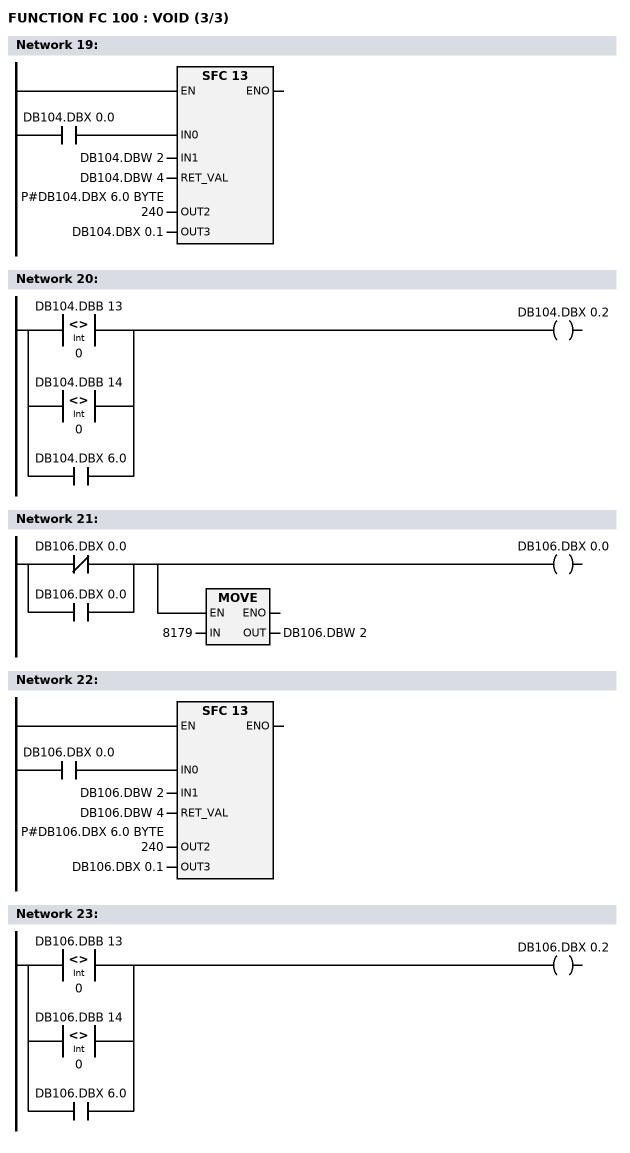

      A     DB104.DBX    0.0;
      =     L      0.0;
      BLD   103;
      CALL SFC   13 (
           IN0                      := L      0.0,
           IN1                      := DB104.DBW    2,
           RET_VAL                  := DB104.DBW    4,
           OUT2                     := P#DB104.DBX 6.0 BYTE 240,
           OUT3                     := DB104.DBX    0.1);
      NOP   0;
NETWORK
TITLE =

      O(    ;
      L     DB104.DBB   13;
      L     0;
      <>I   ;
      )     ;
      O(    ;
      L     DB104.DBB   14;
      L     0;
      <>I   ;
      )     ;
      O     DB104.DBX    6.0;
      =     DB104.DBX    0.2;
NETWORK
TITLE =

      ON    DB106.DBX    0.0;
      O     DB106.DBX    0.0;
      =     L      0.0;
      A     L      0.0;
      BLD   102;
      =     DB106.DBX    0.0;
      A     L      0.0;
      JNB   M003;
      L     8179;
      T     DB106.DBW    2;
M003: NOP   0;
NETWORK
TITLE =

      A     DB106.DBX    0.0;
      =     L      0.0;
      BLD   103;
      CALL SFC   13 (
           IN0                      := L      0.0,
           IN1                      := DB106.DBW    2,
           RET_VAL                  := DB106.DBW    4,
           OUT2                     := P#DB106.DBX 6.0 BYTE 240,
           OUT3                     := DB106.DBX    0.1);
      NOP   0;
NETWORK
TITLE =

      O(    ;
      L     DB106.DBB   13;
      L     0;
      <>I   ;
      )     ;
      O(    ;
      L     DB106.DBB   14;
      L     0;
      <>I   ;
      )     ;
      O     DB106.DBX    6.0;
      =     DB106.DBX    0.2;
END_FUNCTION

DATA_BLOCK DB 500
VERSION : 0.0

 FB 500
BEGIN
   IN0 := FALSE;
   IN1 := FALSE;
   IN2 := FALSE;
   OUT3 := FALSE;
   OUT4 := FALSE;
   STAT5 := FALSE;
   STAT6 := FALSE;
   STAT7 := FALSE;
   STAT8 := FALSE;
END_DATA_BLOCK

DATA_BLOCK DB 501
VERSION : 0.0

 FB 500
BEGIN
   IN0 := FALSE;
   IN1 := FALSE;
   IN2 := FALSE;
   OUT3 := FALSE;
   OUT4 := FALSE;
   STAT5 := FALSE;
   STAT6 := FALSE;
   STAT7 := FALSE;
   STAT8 := FALSE;
END_DATA_BLOCK

DATA_BLOCK DB 502
VERSION : 0.0

 FB 500
BEGIN
   IN0 := FALSE;
   IN1 := FALSE;
   IN2 := FALSE;
   OUT3 := FALSE;
   OUT4 := FALSE;
   STAT5 := FALSE;
   STAT6 := FALSE;
   STAT7 := FALSE;
   STAT8 := FALSE;
END_DATA_BLOCK

DATA_BLOCK DB 504
VERSION : 0.0

 FB 500
BEGIN
   IN0 := FALSE;
   IN1 := FALSE;
   IN2 := FALSE;
   OUT3 := FALSE;
   OUT4 := FALSE;
   STAT5 := FALSE;
   STAT6 := FALSE;
   STAT7 := FALSE;
   STAT8 := FALSE;
END_DATA_BLOCK

DATA_BLOCK DB 505
VERSION : 0.0

 FB 500
BEGIN
   IN0 := FALSE;
   IN1 := FALSE;
   IN2 := FALSE;
   OUT3 := FALSE;
   OUT4 := FALSE;
   STAT5 := FALSE;
   STAT6 := FALSE;
   STAT7 := FALSE;
   STAT8 := FALSE;
END_DATA_BLOCK

DATA_BLOCK DB 506
VERSION : 0.0

 FB 500
BEGIN
   IN0 := FALSE;
   IN1 := FALSE;
   IN2 := FALSE;
   OUT3 := FALSE;
   OUT4 := FALSE;
   STAT5 := FALSE;
   STAT6 := FALSE;
   STAT7 := FALSE;
   STAT8 := FALSE;
END_DATA_BLOCK

DATA_BLOCK DB 507
VERSION : 0.0

 FB 500
BEGIN
   IN0 := FALSE;
   IN1 := FALSE;
   IN2 := FALSE;
   OUT3 := FALSE;
   OUT4 := FALSE;
   STAT5 := FALSE;
   STAT6 := FALSE;
   STAT7 := FALSE;
   STAT8 := FALSE;
END_DATA_BLOCK

DATA_BLOCK DB 508
VERSION : 0.0

 FB 500
BEGIN
   IN0 := FALSE;
   IN1 := FALSE;
   IN2 := FALSE;
   OUT3 := FALSE;
   OUT4 := FALSE;
   STAT5 := FALSE;
   STAT6 := FALSE;
   STAT7 := FALSE;
   STAT8 := FALSE;
END_DATA_BLOCK

DATA_BLOCK DB 509
VERSION : 0.0

 FB 500
BEGIN
   IN0 := FALSE;
   IN1 := FALSE;
   IN2 := FALSE;
   OUT3 := FALSE;
   OUT4 := FALSE;
   STAT5 := FALSE;
   STAT6 := FALSE;
   STAT7 := FALSE;
   STAT8 := FALSE;
END_DATA_BLOCK

DATA_BLOCK DB 512
VERSION : 0.0

 FB 500
BEGIN
   IN0 := FALSE;
   IN1 := FALSE;
   IN2 := FALSE;
   OUT3 := FALSE;
   OUT4 := FALSE;
   STAT5 := FALSE;
   STAT6 := FALSE;
   STAT7 := FALSE;
   STAT8 := FALSE;
END_DATA_BLOCK

DATA_BLOCK DB 516
VERSION : 0.0

 FB 500
BEGIN
   IN0 := FALSE;
   IN1 := FALSE;
   IN2 := FALSE;
   OUT3 := FALSE;
   OUT4 := FALSE;
   STAT5 := FALSE;
   STAT6 := FALSE;
   STAT7 := FALSE;
   STAT8 := FALSE;
END_DATA_BLOCK

DATA_BLOCK DB 517
VERSION : 0.0

 FB 500
BEGIN
   IN0 := FALSE;
   IN1 := FALSE;
   IN2 := FALSE;
   OUT3 := FALSE;
   OUT4 := FALSE;
   STAT5 := FALSE;
   STAT6 := FALSE;
   STAT7 := FALSE;
   STAT8 := FALSE;
END_DATA_BLOCK

DATA_BLOCK DB 518
VERSION : 0.0

 FB 500
BEGIN
   IN0 := FALSE;
   IN1 := FALSE;
   IN2 := FALSE;
   OUT3 := FALSE;
   OUT4 := FALSE;
   STAT5 := FALSE;
   STAT6 := FALSE;
   STAT7 := FALSE;
   STAT8 := FALSE;
END_DATA_BLOCK

DATA_BLOCK DB 520
VERSION : 0.0

 FB 500
BEGIN
   IN0 := FALSE;
   IN1 := FALSE;
   IN2 := FALSE;
   OUT3 := FALSE;
   OUT4 := FALSE;
   STAT5 := FALSE;
   STAT6 := FALSE;
   STAT7 := FALSE;
   STAT8 := FALSE;
END_DATA_BLOCK

DATA_BLOCK DB 521
VERSION : 0.0

 FB 500
BEGIN
   IN0 := FALSE;
   IN1 := FALSE;
   IN2 := FALSE;
   OUT3 := FALSE;
   OUT4 := FALSE;
   STAT5 := FALSE;
   STAT6 := FALSE;
   STAT7 := FALSE;
   STAT8 := FALSE;
END_DATA_BLOCK

DATA_BLOCK DB 522
VERSION : 0.0

 FB 500
BEGIN
   IN0 := FALSE;
   IN1 := FALSE;
   IN2 := FALSE;
   OUT3 := FALSE;
   OUT4 := FALSE;
   STAT5 := FALSE;
   STAT6 := FALSE;
   STAT7 := FALSE;
   STAT8 := FALSE;
END_DATA_BLOCK

DATA_BLOCK DB 523
VERSION : 0.0

 FB 500
BEGIN
   IN0 := FALSE;
   IN1 := FALSE;
   IN2 := FALSE;
   OUT3 := FALSE;
   OUT4 := FALSE;
   STAT5 := FALSE;
   STAT6 := FALSE;
   STAT7 := FALSE;
   STAT8 := FALSE;
END_DATA_BLOCK

DATA_BLOCK DB 525
VERSION : 0.0

 FB 500
BEGIN
   IN0 := FALSE;
   IN1 := FALSE;
   IN2 := FALSE;
   OUT3 := FALSE;
   OUT4 := FALSE;
   STAT5 := FALSE;
   STAT6 := FALSE;
   STAT7 := FALSE;
   STAT8 := FALSE;
END_DATA_BLOCK

DATA_BLOCK DB 526
VERSION : 0.0

 FB 500
BEGIN
   IN0 := FALSE;
   IN1 := FALSE;
   IN2 := FALSE;
   OUT3 := FALSE;
   OUT4 := FALSE;
   STAT5 := FALSE;
   STAT6 := FALSE;
   STAT7 := FALSE;
   STAT8 := FALSE;
END_DATA_BLOCK

DATA_BLOCK DB 527
VERSION : 0.0

 FB 500
BEGIN
   IN0 := FALSE;
   IN1 := FALSE;
   IN2 := FALSE;
   OUT3 := FALSE;
   OUT4 := FALSE;
   STAT5 := FALSE;
   STAT6 := FALSE;
   STAT7 := FALSE;
   STAT8 := FALSE;
END_DATA_BLOCK

DATA_BLOCK DB 528
VERSION : 0.0

 FB 500
BEGIN
   IN0 := FALSE;
   IN1 := FALSE;
   IN2 := FALSE;
   OUT3 := FALSE;
   OUT4 := FALSE;
   STAT5 := FALSE;
   STAT6 := FALSE;
   STAT7 := FALSE;
   STAT8 := FALSE;
END_DATA_BLOCK

DATA_BLOCK DB 529
VERSION : 0.0

 FB 500
BEGIN
   IN0 := FALSE;
   IN1 := FALSE;
   IN2 := FALSE;
   OUT3 := FALSE;
   OUT4 := FALSE;
   STAT5 := FALSE;
   STAT6 := FALSE;
   STAT7 := FALSE;
   STAT8 := FALSE;
END_DATA_BLOCK

DATA_BLOCK DB 530
VERSION : 0.0

 FB 500
BEGIN
   IN0 := FALSE;
   IN1 := FALSE;
   IN2 := FALSE;
   OUT3 := FALSE;
   OUT4 := FALSE;
   STAT5 := FALSE;
   STAT6 := FALSE;
   STAT7 := FALSE;
   STAT8 := FALSE;
END_DATA_BLOCK

DATA_BLOCK DB 531
VERSION : 0.0

 FB 500
BEGIN
   IN0 := FALSE;
   IN1 := FALSE;
   IN2 := FALSE;
   OUT3 := FALSE;
   OUT4 := FALSE;
   STAT5 := FALSE;
   STAT6 := FALSE;
   STAT7 := FALSE;
   STAT8 := FALSE;
END_DATA_BLOCK

DATA_BLOCK DB 532
VERSION : 0.0

 FB 500
BEGIN
   IN0 := FALSE;
   IN1 := FALSE;
   IN2 := FALSE;
   OUT3 := FALSE;
   OUT4 := FALSE;
   STAT5 := FALSE;
   STAT6 := FALSE;
   STAT7 := FALSE;
   STAT8 := FALSE;
END_DATA_BLOCK

DATA_BLOCK DB 534
VERSION : 0.0

 FB 500
BEGIN
   IN0 := FALSE;
   IN1 := FALSE;
   IN2 := FALSE;
   OUT3 := FALSE;
   OUT4 := FALSE;
   STAT5 := FALSE;
   STAT6 := FALSE;
   STAT7 := FALSE;
   STAT8 := FALSE;
END_DATA_BLOCK

DATA_BLOCK DB 535
VERSION : 0.0

 FB 500
BEGIN
   IN0 := FALSE;
   IN1 := FALSE;
   IN2 := FALSE;
   OUT3 := FALSE;
   OUT4 := FALSE;
   STAT5 := FALSE;
   STAT6 := FALSE;
   STAT7 := FALSE;
   STAT8 := FALSE;
END_DATA_BLOCK

DATA_BLOCK DB 510
VERSION : 0.0

 FB 500
BEGIN
   IN0 := FALSE;
   IN1 := FALSE;
   IN2 := FALSE;
   OUT3 := FALSE;
   OUT4 := FALSE;
   STAT5 := FALSE;
   STAT6 := FALSE;
   STAT7 := FALSE;
   STAT8 := FALSE;
END_DATA_BLOCK

DATA_BLOCK DB 511
VERSION : 0.0

 FB 500
BEGIN
   IN0 := FALSE;
   IN1 := FALSE;
   IN2 := FALSE;
   OUT3 := FALSE;
   OUT4 := FALSE;
   STAT5 := FALSE;
   STAT6 := FALSE;
   STAT7 := FALSE;
   STAT8 := FALSE;
END_DATA_BLOCK

DATA_BLOCK DB 513
VERSION : 0.0

 FB 500
BEGIN
   IN0 := FALSE;
   IN1 := FALSE;
   IN2 := FALSE;
   OUT3 := FALSE;
   OUT4 := FALSE;
   STAT5 := FALSE;
   STAT6 := FALSE;
   STAT7 := FALSE;
   STAT8 := FALSE;
END_DATA_BLOCK

DATA_BLOCK DB 514
VERSION : 0.0

 FB 500
BEGIN
   IN0 := FALSE;
   IN1 := FALSE;
   IN2 := FALSE;
   OUT3 := FALSE;
   OUT4 := FALSE;
   STAT5 := FALSE;
   STAT6 := FALSE;
   STAT7 := FALSE;
   STAT8 := FALSE;
END_DATA_BLOCK

DATA_BLOCK DB 515
VERSION : 0.0

 FB 500
BEGIN
   IN0 := FALSE;
   IN1 := FALSE;
   IN2 := FALSE;
   OUT3 := FALSE;
   OUT4 := FALSE;
   STAT5 := FALSE;
   STAT6 := FALSE;
   STAT7 := FALSE;
   STAT8 := FALSE;
END_DATA_BLOCK

DATA_BLOCK DB 519
VERSION : 0.0

 FB 500
BEGIN
   IN0 := FALSE;
   IN1 := FALSE;
   IN2 := FALSE;
   OUT3 := FALSE;
   OUT4 := FALSE;
   STAT5 := FALSE;
   STAT6 := FALSE;
   STAT7 := FALSE;
   STAT8 := FALSE;
END_DATA_BLOCK

DATA_BLOCK DB 524
VERSION : 0.0

 FB 500
BEGIN
   IN0 := FALSE;
   IN1 := FALSE;
   IN2 := FALSE;
   OUT3 := FALSE;
   OUT4 := FALSE;
   STAT5 := FALSE;
   STAT6 := FALSE;
   STAT7 := FALSE;
   STAT8 := FALSE;
END_DATA_BLOCK

DATA_BLOCK DB 533
VERSION : 0.0

 FB 500
BEGIN
   IN0 := FALSE;
   IN1 := FALSE;
   IN2 := FALSE;
   OUT3 := FALSE;
   OUT4 := FALSE;
   STAT5 := FALSE;
   STAT6 := FALSE;
   STAT7 := FALSE;
   STAT8 := FALSE;
END_DATA_BLOCK

ORGANIZATION_BLOCK OB 1
VERSION : 0.1


VAR_TEMP
  TEMP0 : BYTE ;
  TEMP1 : BYTE ;
  TEMP2 : BYTE ;
  TEMP3 : BYTE ;
  TEMP4 : BYTE ;
  TEMP5 : BYTE ;
  TEMP6 : INT ;
  TEMP7 : INT ;
  TEMP8 : INT ;
  TEMP9 : DATE_AND_TIME ;
END_VAR
BEGIN
NETWORK
TITLE =
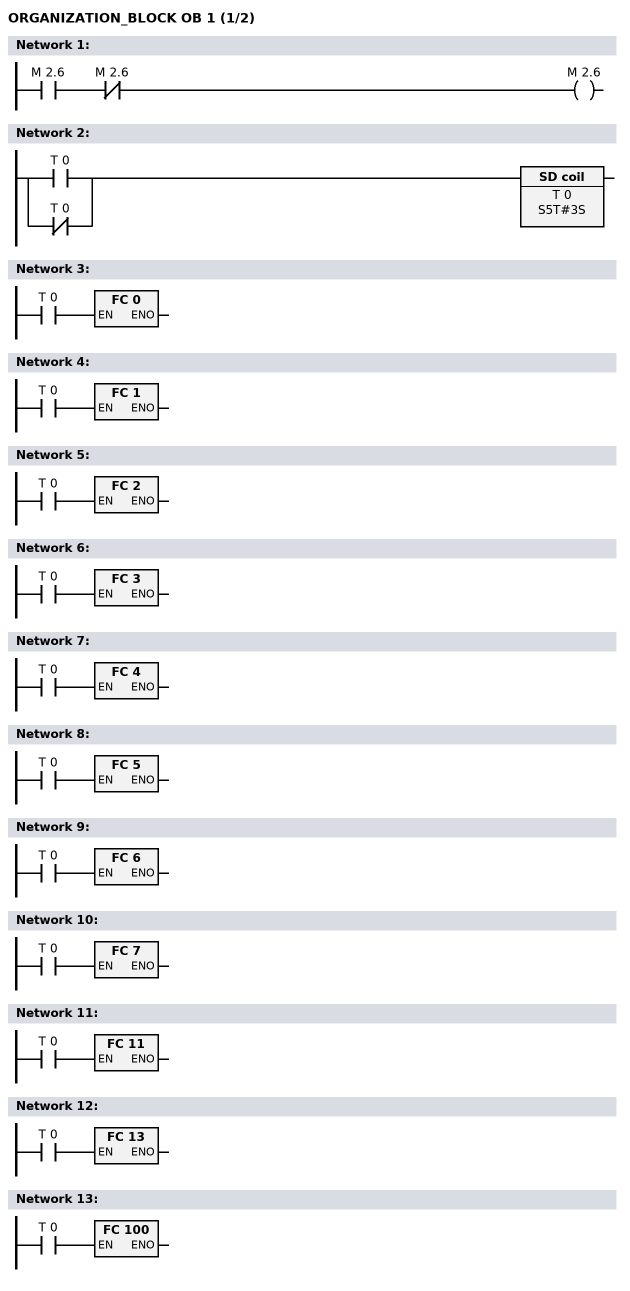

      A     M      2.6;
      AN    M      2.6;
      =     M      2.6;
NETWORK
TITLE =

      A(    ;
      O     T      0;
      ON    T      0;
      )     ;
      L     S5T#3S;
      SD    T      0;
      NOP   0;
      NOP   0;
      NOP   0;
      NOP   0;
NETWORK
TITLE =

      A     T      0;
      JNB   M001;
      CALL FC     0 ;
M001: NOP   0;
NETWORK
TITLE =

      A     T      0;
      JNB   M002;
      CALL FC     1 ;
M002: NOP   0;
NETWORK
TITLE =

      A     T      0;
      JNB   M003;
      CALL FC     2 ;
M003: NOP   0;
NETWORK
TITLE =

      A     T      0;
      JNB   M004;
      CALL FC     3 ;
M004: NOP   0;
NETWORK
TITLE =

      A     T      0;
      JNB   M005;
      CALL FC     4 ;
M005: NOP   0;
NETWORK
TITLE =

      A     T      0;
      JNB   M006;
      CALL FC     5 ;
M006: NOP   0;
NETWORK
TITLE =

      A     T      0;
      JNB   M007;
      CALL FC     6 ;
M007: NOP   0;
NETWORK
TITLE =

      A     T      0;
      JNB   M008;
      CALL FC     7 ;
M008: NOP   0;
NETWORK
TITLE =

      A     T      0;
      JNB   M009;
      CALL FC    11 ;
M009: NOP   0;
NETWORK
TITLE =

      A     T      0;
      JNB   M00a;
      CALL FC    13 ;
M00a: NOP   0;
NETWORK
TITLE =

      A     T      0;
      JNB   M00b;
      CALL FC   100 ;
M00b: NOP   0;
NETWORK
TITLE =
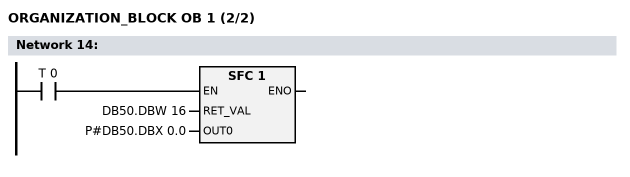

      A     T      0;
      JNB   M00c;
      CALL SFC    1 (
           RET_VAL                  := DB50.DBW   16,
           OUT0                     := P#DB50.DBX 0.0);
M00c: NOP   0;
END_ORGANIZATION_BLOCK

ORGANIZATION_BLOCK OB 35
VERSION : 0.1


VAR_TEMP
  TEMP0 : BYTE ;
  TEMP1 : BYTE ;
  TEMP2 : BYTE ;
  TEMP3 : BYTE ;
  TEMP4 : BYTE ;
  TEMP5 : BYTE ;
  TEMP6 : WORD ;
  TEMP7 : INT ;
  TEMP8 : INT ;
  TEMP9 : DATE_AND_TIME ;
END_VAR
BEGIN
END_ORGANIZATION_BLOCK

ORGANIZATION_BLOCK OB 70
VERSION : 0.1


VAR_TEMP
  TEMP0 : BYTE ;
  TEMP1 : BYTE ;
  TEMP2 : BYTE ;
  TEMP3 : BYTE ;
  TEMP4 : WORD ;
  TEMP5 : WORD ;
  TEMP6 : WORD ;
  TEMP7 : WORD ;
  TEMP8 : DATE_AND_TIME ;
END_VAR
BEGIN
NETWORK
TITLE =

      AN    M      3.7;
      =     M      3.7;
END_ORGANIZATION_BLOCK

ORGANIZATION_BLOCK OB 72
VERSION : 0.1


VAR_TEMP
  TEMP0 : BYTE ;
  TEMP1 : BYTE ;
  TEMP2 : BYTE ;
  TEMP3 : BYTE ;
  TEMP4 : WORD ;
  TEMP5 : WORD ;
  TEMP6 : WORD ;
  TEMP7 : WORD ;
  TEMP8 : DATE_AND_TIME ;
END_VAR
BEGIN
NETWORK
TITLE =

      A     M      3.7;
      =     M      3.7;
END_ORGANIZATION_BLOCK

ORGANIZATION_BLOCK OB 81
VERSION : 0.1


VAR_TEMP
  TEMP0 : BYTE ;
  TEMP1 : BYTE ;
  TEMP2 : BYTE ;
  TEMP3 : BYTE ;
  TEMP4 : BYTE ;
  TEMP5 : BYTE ;
  TEMP6 : WORD ;
  TEMP7 : BYTE ;
  TEMP8 : BYTE ;
  TEMP9 : BYTE ;
  TEMP10 : BYTE ;
  TEMP11 : DATE_AND_TIME ;
END_VAR
BEGIN
NETWORK
TITLE =

      AN    M      3.7;
      =     M      3.7;
END_ORGANIZATION_BLOCK

ORGANIZATION_BLOCK OB 82
VERSION : 0.1


VAR_TEMP
  TEMP0 : BYTE ;
  TEMP1 : BYTE ;
  TEMP2 : BYTE ;
  TEMP3 : BYTE ;
  TEMP4 : BYTE ;
  TEMP5 : BYTE ;
  TEMP6 : WORD ;
  TEMP7 : BOOL ;
  TEMP8 : BOOL ;
  TEMP9 : BOOL ;
  TEMP10 : BOOL ;
  TEMP11 : BOOL ;
  TEMP12 : BOOL ;
  TEMP13 : BOOL ;
  TEMP14 : BOOL ;
  TEMP15 : BYTE ;
  TEMP16 : BOOL ;
  TEMP17 : BOOL ;
  TEMP18 : BOOL ;
  TEMP19 : BOOL ;
  TEMP20 : BOOL ;
  TEMP21 : BOOL ;
  TEMP22 : BOOL ;
  TEMP23 : BOOL ;
  TEMP24 : BOOL ;
  TEMP25 : BOOL ;
  TEMP26 : BOOL ;
  TEMP27 : BOOL ;
  TEMP28 : BOOL ;
  TEMP29 : BOOL ;
  TEMP30 : BOOL ;
  TEMP31 : BOOL ;
  TEMP32 : DATE_AND_TIME ;
END_VAR
BEGIN
NETWORK
TITLE =

      AN    M      3.7;
      =     M      3.7;
END_ORGANIZATION_BLOCK

ORGANIZATION_BLOCK OB 83
VERSION : 0.1


VAR_TEMP
  TEMP0 : BYTE ;
  TEMP1 : BYTE ;
  TEMP2 : BYTE ;
  TEMP3 : BYTE ;
  TEMP4 : BYTE ;
  TEMP5 : BYTE ;
  TEMP6 : WORD ;
  TEMP7 : INT ;
  TEMP8 : WORD ;
  TEMP9 : DATE_AND_TIME ;
END_VAR
BEGIN
NETWORK
TITLE =

      AN    M      3.7;
      =     M      3.7;
END_ORGANIZATION_BLOCK

ORGANIZATION_BLOCK OB 85
VERSION : 0.1


VAR_TEMP
  TEMP0 : BYTE ;
  TEMP1 : BYTE ;
  TEMP2 : BYTE ;
  TEMP3 : BYTE ;
  TEMP4 : BYTE ;
  TEMP5 : BYTE ;
  TEMP6 : INT ;
  TEMP7 : BYTE ;
  TEMP8 : BYTE ;
  TEMP9 : BYTE ;
  TEMP10 : BYTE ;
  TEMP11 : DATE_AND_TIME ;
END_VAR
BEGIN
NETWORK
TITLE =

      AN    M      3.7;
      =     M      3.7;
END_ORGANIZATION_BLOCK

ORGANIZATION_BLOCK OB 86
VERSION : 0.1


VAR_TEMP
  TEMP0 : BYTE ;
  TEMP1 : BYTE ;
  TEMP2 : BYTE ;
  TEMP3 : BYTE ;
  TEMP4 : BYTE ;
  TEMP5 : BYTE ;
  TEMP6 : WORD ;
  TEMP7 : ARRAY  [0 .. 31 ] OF BOOL ;
  TEMP8 : DATE_AND_TIME ;
END_VAR
BEGIN
NETWORK
TITLE =

      AN    M      3.7;
      =     M      3.7;
END_ORGANIZATION_BLOCK

ORGANIZATION_BLOCK OB 87
VERSION : 0.1


VAR_TEMP
  TEMP0 : BYTE ;
  TEMP1 : BYTE ;
  TEMP2 : BYTE ;
  TEMP3 : BYTE ;
  TEMP4 : BYTE ;
  TEMP5 : BYTE ;
  TEMP6 : WORD ;
  TEMP7 : DWORD ;
  TEMP8 : DATE_AND_TIME ;
END_VAR
BEGIN
NETWORK
TITLE =

      AN    M      3.7;
      =     M      3.7;
END_ORGANIZATION_BLOCK

ORGANIZATION_BLOCK OB 100
VERSION : 0.1


VAR_TEMP
  TEMP0 : BYTE ;
  TEMP1 : BYTE ;
  TEMP2 : BYTE ;
  TEMP3 : BYTE ;
  TEMP4 : BYTE ;
  TEMP5 : BYTE ;
  TEMP6 : WORD ;
  TEMP7 : DWORD ;
  TEMP8 : DATE_AND_TIME ;
END_VAR
BEGIN
END_ORGANIZATION_BLOCK

ORGANIZATION_BLOCK OB 122
VERSION : 0.1


VAR_TEMP
  TEMP0 : BYTE ;
  TEMP1 : BYTE ;
  TEMP2 : BYTE ;
  TEMP3 : BYTE ;
  TEMP4 : BYTE ;
  TEMP5 : BYTE ;
  TEMP6 : WORD ;
  TEMP7 : WORD ;
  TEMP8 : WORD ;
  TEMP9 : DATE_AND_TIME ;
END_VAR
BEGIN
NETWORK
TITLE =

      AN    M      3.7;
      =     M      3.7;
END_ORGANIZATION_BLOCK

